(* IEC 61131-3 sources: plc-iiot-stack/src/POUs/Iiot/F_IiotIsPrintable, 2 files *)

(* ---- F_IiotIsPrintable.decl.st ---- *)
// Назначение: строка из печатных символов ASCII (пробел..~) длиной 1..iMaxLen (поле origin).
// Автор:      kr0nsch
// Версия:     0.1.0
// Документ:   docs/plc_mqtt.md, раздел «Команды»
FUNCTION F_IiotIsPrintable : BOOL
VAR_INPUT
    sText : STRING(GVL_Const.JSON_STR_LEN);
    iMaxLen : INT;
END_VAR
VAR
    iLen : INT;
    iIdx : INT;
    bCh : BYTE;
END_VAR

(* ---- F_IiotIsPrintable.impl.st ---- *)
iLen := LEN(sText);
IF iLen < 1 OR iLen > iMaxLen THEN
    RETURN;
END_IF
FOR iIdx := 0 TO iLen - 1 DO
    bCh := sText[iIdx];
    IF bCh < GVL_Const.ASCII_SPACE OR bCh > GVL_Const.ASCII_TILDE THEN
        RETURN;
    END_IF
END_FOR
F_IiotIsPrintable := TRUE;
